// TIA Portal V19 export
DATA_BLOCK "Tacho2_UM"   // DB1
VERSION : 1.0
// stored: InstanceOfName UM_Principal, InstanceOfType FB
"UM_Principal"
   // VAR_INPUT
   //    UM_Ctrl : "EM_Input";
   //    Recipe : Int;
   //    SelMeladura : Int;
   //    NivelTacho : Real;
   //    SobreSaturacion : Real;
   //    ControlExtOk : Bool;
   //    ConcSMMV : Real;
   //    VaccumSMMV : Real;
   //    FeedSMMV : Real;
   //    EM01_Estado : "EM01_Output";
   //    EM02_Estado : "EM02_Output";
   //    EM03_Estado : "EM03_Output";
   //    EM04_Estado : "EM04_Output";
   //    EM05_Estado : "EM05_Output";
   //    EM06_Estado : "EM06_Output";
   //    ParametrosDeControlGeneral : Struct
   //       SPTemperaturaCalentamiento : Real;
   //       TimeoutCalentamiento : Time;
   //       SPVacioCuerpo : Real;
   //       TimeoutVacio : Time;
   //       BandaVacio : Real;
   //       SPConcentracionStrike : Real;
   //       BandaConcentracion : Real;
   //       TiempoEstabConcentracion : Time;
   //       PosicionHoldCalandria : Real;
   //       NivelRunAgitador : Real;
   //       NivelAbrirDescarga : Real;
   //       NivelCerrarDescarga : Real;
   //       NivelFinDescarga : Real;
   //       PurezaSemilla : Real;
   //       PurezaCorte : Real;
   //       PurezasInsumos : Array[1..2] of Real;
   //    END_STRUCT;
   //    ParametrosDeControlSlurry : Struct
   //       SPNivelPieInicial : Real;
   //       SP_SS_Preaviso : Real;
   //       SP_SS_Siembra : Real;
   //       SP_TiempoSiembra : Time;
   //       SP_TiempoMaduracion : Time;
   //       SP_Nivel_Final_Coccion : Real;
   //       SP_Brix_Final_Coccion : Real;
   //       SP_Brix_Final_Secado : Real;
   //       SP_VacioPausa : Real;
   //    END_STRUCT;
   //    BrixMasaActual : Real;
   //    BrixLicorActual : Real;
   // END_VAR
   // VAR_OUTPUT
   //    UM_State : "EM_Output";
   //    Seed_Advice : Bool;
   //    ExternalControlCmds : Struct
   //       Purity_P1 : Real;
   //       Purity_P2 : Real;
   //       Purity_P3 : Real;
   //       Purity_Selector : UInt;
   //       Final_Mass_Solid_Prog1 : Real;
   //       Final_Mass_Solid_Prog2 : Real;
   //       Final_Mass_Solid_Prog3 : Real;
   //       Final_Mass_Solid_Selector : UInt;
   //       Strike_Active : Bool;
   //       Seeded : Bool;
   //    END_STRUCT;
   //    EM01_Comandos : "EM01_Input";
   //    EM02_Comandos : "EM02_Input";
   //    EM03_Comandos : "EM03_Input";
   //    EM04_Comandos : "EM04_Input";
   //    EM05_Comandos : "EM05_Input";
   //    EM06_Comandos : "EM06_Input";
   // END_VAR
   // VAR
   //    State : Int;
   //    "Step" : Int;
   //    RecipeActiva : Int;
   //    MeladuraActiva : Int;
   //    ConfigFault : Int;
   //    NivelAgitadorOk : Bool;
   //    StartEM05Prev : Bool;
   //    SeedStartIssued : Bool;
   //    MaturationElapsed : Time;
   //    ModoExt : Bool;
   //    NivelCocicionInicial : Real;
   //    BrixMasaInicial : Real;
   //    BrixLicorInicial : Real;
   //    CocicionEnPausa : Bool;
   //    ModoExtCocicion : Bool;
   //    TimerMaduracion { S7_SetPoint := 'True'} : TON_TIME;
   //    TrigStart { S7_SetPoint := 'True'} : R_TRIG;
   //    TrigStop { S7_SetPoint := 'True'} : R_TRIG;
   //    TrigHold { S7_SetPoint := 'True'} : R_TRIG;
   //    TrigAbort { S7_SetPoint := 'True'} : R_TRIG;
   //    TrigReset { S7_SetPoint := 'True'} : R_TRIG;
   //    PurezaP1_Value : Real;
   //    PurezaP2_Value : Real;
   //    PurezaP3_Value : Real;
   //    PurezasValoresLatcheadas : Bool;
   // END_VAR
BEGIN
END_DATA_BLOCK
